(* IEC 61131-3 sources: volt/packages/volt-lsp-iec/test-corpus/bakon-nano/Device/Plc Logic/Application/Library Manager/AlarmManager (part 4) *)

(* ---- STANDARDALARMCONFIGURATION.pou ---- *)
FUNCTION_BLOCK STANDARDALARMCONFIGURATION
VAR
	M_PAITFALARMGROUPS : POINTER TO ARRAY [0..0] OF IAlarmGroup;
	M_ICOUNTALARMGROUPS : INT;
	M_PAITFALARMCLASSES : POINTER TO ARRAY [0..0] OF IAlarmClass;
	M_ICOUNTALARMCLASSES : INT;
	M_XVARIABLESREGISTERED : BOOL;
	M_XFIRST : BOOL;
	M_XPLACEHOLDANALYZED : BOOL;
	M_LTSTARTTIME : LTIME;
	M_DATABASESIZELIMIT : DatabaseSizeLimit;
	M_XDATABASESIZELIMITBLOCKED : BOOL;
	_XRAISEDMOREALARMSTHANSTORAGELIMITREPORTED : BOOL;
	_XCLEARHISTORY : BOOL;
	_XKEEPACTIVEALARMS : BOOL;
	M_DICTALARMTEMPLATEINSTANCES : AlarmInstanceDictionary;
	M_SZAPPNAME : STRING(CmpApp.GlobalConstants.MAX_LEN_APPLNAME);
	DATABASESIZELIMIT : IDatabaseSizeLimit;
	TOTALROWSTOINSERT : UDINT;
END_VAR
END_FUNCTION_BLOCK

METHOD FB_EXIT : BOOL
VAR_INPUT
	BINCOPYCODE : BOOL;
END_VAR
END_METHOD

METHOD FB_INIT : BOOL
VAR_INPUT
	BINITRETAINS : BOOL;
	BINCOPYCODE : BOOL;
END_VAR
END_METHOD

METHOD FINDALARMBYID : IAlarm
VAR_INPUT
	USIALARMGROUPID : ALARMGROUP_ID;
	UIALARMID : ALARM_ID;
END_VAR
END_METHOD

METHOD REGISTERVARIABLES
END_METHOD

METHOD ADDTOINSTANCEDICTIONARY : BOOL
VAR_INPUT
	PINSTANCE : POINTER TO BYTE;
	PSTALARMTEMPLATENAME : POINTER TO STRING;
	UDIALARMGROUPID : UDINT;
	UITEMPLATEALARMSOFFSET : UINT;
	UITEMPLATEALARMSLENGTH : UINT;
	UITEMPLATEEVENTSOFFSET : UINT;
	UITEMPLATEEVENTSLENGTH : UINT;
END_VAR
END_METHOD

METHOD CLEARINSTANCEDICTIONARY : BOOL
END_METHOD

METHOD GETALARMFROMDICTIONARY : IAlarm8
VAR_INPUT
	PINSTANCE : POINTER TO BYTE;
	UDIALARMID : REFERENCE TO ALARM_ID;
	STALARMTEMPLATENAME : REFERENCE TO STRING;
END_VAR
VAR_OUTPUT
	USIALARMGROUPID : ALARMGROUP_ID;
	UIALARMID : ALARM_ID;
END_VAR
END_METHOD

METHOD CREATEALARMSTORAGETASK
VAR_INPUT
	STSTORAGETASKGROUPNAME : REFERENCE TO STRING;
END_VAR
END_METHOD

METHOD INITSTORAGETASKINFO
VAR_INPUT
	ITASKPRIORITY : INT;
	DWINTERVAL : DWORD;
END_VAR
END_METHOD

METHOD ACKNOWLEDGEALL
END_METHOD

METHOD ACKNOWLEDGEALLOFGROUP
VAR_INPUT
	USIALARMGROUPID : ALARMGROUP_ID;
END_VAR
END_METHOD

METHOD ACKNOWLEDGEONEOFGROUP
VAR_INPUT
	USIALARMGROUPID : ALARMGROUP_ID;
	UIALARMID : ALARM_ID;
END_VAR
END_METHOD

METHOD CYCLICCALL
END_METHOD

METHOD FINDALARM : POINTER TO Alarm
VAR_INPUT
	SALARMGROUP : STRING;
	UIALARMID : ALARM_ID;
END_VAR
END_METHOD

METHOD FINDALARMCLASS : IAlarmClass
VAR_INPUT
	UDIID : UDINT;
END_VAR
END_METHOD

METHOD FINDALARMGROUP : IAlarmGroup
VAR_INPUT
	UDIID : UDINT;
END_VAR
END_METHOD

METHOD GETSTORAGE : IDatabaseFileAlarmStorage
END_METHOD

METHOD HASSTORAGE : BOOL
END_METHOD

METHOD RAISEEVENT : BOOL
VAR_INPUT
	EVENT : AlarmEvent;
END_VAR
END_METHOD

METHOD DETERMINERELEVANTALARMS : UDINT
VAR_INPUT
	ITFALARMFILTERCRITERIA : IAlarmFilterCriteria;
	PARRITFRELEVANTALARMS : POINTER TO ARRAY [0..0] OF IAlarm;
	IOFFSET : INT;
END_VAR
END_METHOD

METHOD FINDALARMGROUPBYNAME : IAlarmGroup
VAR_INPUT
	SALARMGROUP : STRING;
END_VAR
END_METHOD

METHOD FINDALARMCLASSBYNAME : IAlarmClass
VAR_INPUT
	SALARMCLASS : STRING;
END_VAR
END_METHOD

METHOD RAISEEVENT2 : BOOL
VAR_INPUT
	EVENT : AlarmEvent;
END_VAR
VAR_OUTPUT
	ITFALARM : IAlarm;
END_VAR
END_METHOD

METHOD GETALARMGROUPS : POINTER TO ARRAY [0..0] OF IAlarmGroup
VAR_OUTPUT
	IALARMGROUPCOUNT : INT;
END_VAR
END_METHOD

METHOD FINDALARMCLASSCOUNT : INT
END_METHOD

METHOD CLEARHISTORY : BOOL
VAR_INPUT
	XKEEPACTIVEALARMS : BOOL;
END_VAR
END_METHOD

METHOD ACKNOWLEDGEALLOFGROUPWITHCOMMENT
VAR_INPUT
	USIALARMGROUPID : ALARMGROUP_ID;
END_VAR
VAR_IN_OUT
	WSCOMMENT : WSTRING;
	WSUSERID : WSTRING;
END_VAR
END_METHOD

METHOD ACKNOWLEDGEALLWITHCOMMENT
VAR_IN_OUT
	WSCOMMENT : WSTRING;
	WSUSERID : WSTRING;
END_VAR
END_METHOD

METHOD ACKNOWLEDGEONEOFGROUPWITHCOMMENT
VAR_INPUT
	USIALARMGROUPID : ALARMGROUP_ID;
	UIALARMID : ALARM_ID;
END_VAR
VAR_IN_OUT
	WSCOMMENT : WSTRING;
	WSUSERID : WSTRING;
END_VAR
END_METHOD

METHOD SETCOMMENT : UDINT
VAR_INPUT
	USIALARMGROUPID : ALARMGROUP_ID;
	UIALARMID : ALARM_ID;
END_VAR
VAR_IN_OUT
	WSCOMMENT : WSTRING;
	WSUSERID : WSTRING;
END_VAR
END_METHOD

METHOD TRAVERSEALLALARMSOFALLALARMGROUPS
VAR_INPUT
	ITFALARMTRAVERSALCONSUMER : IAlarmTraversalConsumer;
END_VAR
END_METHOD

METHOD TRAVERSEALLCLASSES
VAR_INPUT
	ITFALARMTRAVERSALCONSUMER : IAlarmTraversalConsumer;
END_VAR
END_METHOD

METHOD NOTIFYREINITDONE
END_METHOD

METHOD CLEARALLALARMHISTORYENTRIESIFWISHED : BOOL
VAR_INPUT
	ITFDATABASEFILEALARMSTORAGE : IDatabaseFileAlarmStorage;
END_VAR
END_METHOD

METHOD CLEARONLYHISTORYOFINACTIVEALARMS : BOOL
END_METHOD

METHOD PRVACKNOWLEDGE
VAR_INPUT
	PAALARMS : POINTER TO ARRAY [0..0] OF Alarm;
	IALARMCOUNT : INT;
	UIALARMID : ALARM_ID;
	XACKALL : BOOL;
	PWSCOMMENT : POINTER TO WSTRING;
	PWSUSER : POINTER TO WSTRING;
END_VAR
END_METHOD

METHOD PRVCHECKSETACKNOWLEDGE
VAR_INPUT
	INDEX : INT;
	UIALARMID : ALARM_ID;
	XACKALL : BOOL;
	PWSCOMMENT : POINTER TO WSTRING;
	PWSUSER : POINTER TO WSTRING;
END_VAR
END_METHOD

METHOD PRVCREATEALARMSTORAGEMETADATAFILE
END_METHOD

METHOD PRVDETERMINERELEVANTALARMS : UDINT
VAR_INPUT
	PAALARMS : POINTER TO ARRAY [0..0] OF Alarm;
	IALARMCOUNT : INT;
	ITFALARMFILTERCRITERIA : IAlarmFilterCriteria;
	PARRITFRELEVANTALARMS : POINTER TO ARRAY [0..0] OF IAlarm;
	IOFFSET : INT;
END_VAR
END_METHOD

METHOD PRVINITIALIZEALARMCONFIGURATION
END_METHOD

METHOD PRVTRYGETCURRENTROW : BOOL
VAR_OUTPUT
	CURRENTROW : AlarmStorageRow;
END_VAR
END_METHOD

METHOD PRVTSTPLACEHOLDERS : BOOL
VAR_INPUT
	ALARM : REFERENCE TO Alarm;
END_VAR
END_METHOD

METHOD PRVWITHBRACKETS : STRING
VAR_INPUT
	SSTRING : STRING;
END_VAR
END_METHOD

METHOD PRVWITHOPENINGBRACKET : STRING
VAR_INPUT
	SSTRING : STRING;
END_VAR
END_METHOD

(* ---- STANDARDALARMCONFIGURATIONREMOTE.pou ---- *)
FUNCTION_BLOCK STANDARDALARMCONFIGURATIONREMOTE
VAR_INPUT
	M_PAITFPROXY : POINTER TO ARRAY [0..10] OF IProxy;
	M_IPROXYNUM : INT;
END_VAR
VAR
	M_SIALREADYSCAN : SINT := -1;
	PROXYNUM : INT;
END_VAR
END_FUNCTION_BLOCK

METHOD CYCLICCALL
END_METHOD

METHOD GETACTIVEALARMS
VAR_INPUT
	PASNAME : POINTER TO ARRAY [0..10] OF STRING;
	IGROUPCOUNT : INT;
	FILTERCRITERIA : REFERENCE TO VisuFbAlarmFilterCriteria;
	ITFALARMDATABLOCK : IAlarmDataBlockBaseDINT;
END_VAR
VAR_IN_OUT
	DISTUBPROG : DINT;
END_VAR
END_METHOD

METHOD GETALARMCLASSDESC : BOOL
VAR_INPUT
	SPROXYNAME : STRING;
	UDIID : UDINT;
END_VAR
VAR_OUTPUT
	SDESC : ProxyStructAlarmClassDesc;
END_VAR
END_METHOD

METHOD GETALARMCLASSDESCBYNAME : BOOL
VAR_INPUT
	SPROXYNAME : STRING;
	SCLASSNAME : STRING;
END_VAR
VAR_OUTPUT
	SDESC : ProxyStructAlarmClassDesc;
END_VAR
END_METHOD

METHOD GETALARMDESC : BOOL
VAR_INPUT
	SPROXYNAME : STRING;
	UDIALMID : UDINT;
	UDIGRPID : UDINT;
END_VAR
VAR_OUTPUT
	SDESC : ProxyStructAlarmDesc;
END_VAR
END_METHOD

METHOD GETALARMDISPLAYOPTIONS : BOOL
VAR_INPUT
	ITFALARMMETAOBJECTSTUB5 : IAlarmMetaObjectStub5;
	REFDISPLAYOPTIONS : REFERENCE TO DisplayOptions;
END_VAR
VAR_OUTPUT
	XVALID : BOOL;
	SCLASSREMAP : STRING;
END_VAR
END_METHOD

METHOD GETALARMGROUPDESC : BOOL
VAR_INPUT
	SPROXYNAME : STRING;
	UDIID : UDINT;
END_VAR
VAR_OUTPUT
	SDESC : ProxyStructAlarmGroupDesc;
END_VAR
END_METHOD

METHOD GETALARMGROUPDESCBYNAME : BOOL
VAR_INPUT
	SPROXYNAME : STRING;
	SGRPNAME : STRING;
END_VAR
VAR_OUTPUT
	SDESC : ProxyStructAlarmGroupDesc;
END_VAR
END_METHOD

METHOD GETALARMMESSAGE : BOOL
VAR_INPUT
	ITFALARMMETAOBJECTSTUB5 : IAlarmMetaObjectStub5;
	IWHICHMESSAGE : INT;
	REFCHARBUFFERSTRING : REFERENCE TO CharBufferString;
	STRINGTYPE : __SYSTEM.TYPE_CLASS;
END_VAR
END_METHOD

METHOD GETALARMMESSAGE2 : BOOL
VAR_INPUT
	SNAME : STRING;
	STEXTLISTNAME : STRING;
	STEXTLISTINDEX : STRING;
	IWHICHMESSAGE : INT;
	STRINGTYPE : __SYSTEM.TYPE_CLASS;
END_VAR
VAR_OUTPUT
	MESSAGE : CharBufferPtr;
END_VAR
END_METHOD

METHOD GETPROXY : IProxy
VAR_INPUT
	SNAME : STRING;
END_VAR
END_METHOD

METHOD GETSTORAGE : IDatabaseFileAlarmStorage
END_METHOD

METHOD HASSTORAGE : BOOL
END_METHOD

METHOD REGISTERUSERCLIENT : BOOL
VAR_INPUT
	IINDEX : INT;
END_VAR
VAR_OUTPUT
	ITFPROXY : IProxy;
END_VAR
END_METHOD

METHOD SETALARMSTOACK
VAR_INPUT
	ITFALARMDATABLOCK : IAlarmDataBlockBase2;
END_VAR
END_METHOD

METHOD REMOTEDEVICEREACHED
VAR_INPUT
	ROW : REFERENCE TO AlarmStorageRow;
	XFIRST : BOOL;
	IVERSION : INT;
END_VAR
END_METHOD

METHOD PRVGETPROXY : IProxy
VAR_INPUT
	SNAME : STRING;
END_VAR
END_METHOD

METHOD GETPROXYALARMCLASSESDESCRIPTION : BOOL
VAR_INPUT
	SNAME : STRING;
	PCLDESC : POINTER TO ARRAY [0..0] OF ProxyStructMonitorAlarmClassDesc;
	ISIZE : INT;
END_VAR
VAR_OUTPUT
	ICLCNT : INT;
END_VAR
END_METHOD

METHOD GETPROXYALARMGROUPSDESCRIPTION : BOOL
VAR_INPUT
	SNAME : STRING;
	PGRPDESC : POINTER TO ARRAY [0..0] OF ProxyStructMonitorAlarmGroupDesc;
	ISIZE : INT;
END_VAR
VAR_OUTPUT
	IGRPCNT : INT;
END_VAR
END_METHOD

METHOD GETPROXYALARMSDESCRIPTION : BOOL
VAR_INPUT
	SNAME : STRING;
	PALMDESC : POINTER TO ARRAY [0..0] OF ProxyStructMonitorAlarmDesc;
	DISIZE : DINT;
END_VAR
VAR_OUTPUT
	DIALMCNT : DINT;
END_VAR
END_METHOD

METHOD GETPROXYSTATISTICS : BOOL
VAR_INPUT
	SNAME : STRING;
END_VAR
VAR_OUTPUT
	STRUCTMONITOR : ProxyStructMonitor;
END_VAR
END_METHOD

METHOD GETPROXYSTATISTICSSINGLEACTIVITY : BOOL
VAR_INPUT
	SNAME : STRING;
	ITASKID : INT;
END_VAR
VAR_OUTPUT
	STRUCTMONITOR : ProxyStructMonitorRequest;
END_VAR
END_METHOD

(* ---- STANDARDALARMHANDLER.pou ---- *)
FUNCTION_BLOCK STANDARDALARMHANDLER
VAR
	M_AITFALARMCONFIGURATIONS : ARRAY [0..(MAX_COUNT_CONFIG - 1)] OF IAlarmConfiguration;
	M_ICOUNTCONFIGURATIONS : INT := 0;
	M_AITFALARMCONFIGURATIONSREM : ARRAY [0..(MAX_COUNT_CONFIG - 1)] OF IAlarmConfigurationRemote;
	M_ICOUNTCONFIGURATIONSREM : INT := 0;
	M_ALARMMANAGERCLIENTINFOSTRUCTVECTOR : AlarmManagerClientInfoStructVector;
	M_DIALARMSTATETRANSITIONCOUNTERPREVIOUSCALL : DINT;
	M_DIALARMSTORAGECOUNTERPREVIOUSCALL : DINT;
	M_ITFSTORAGETODELETE : IDatabaseFileAlarmStorage;
	M_XSTART : BOOL := TRUE;
	M_XFIRSTCYCLEAFTERDOWNLOAD : BOOL := TRUE;
	MAX_COUNT_CONFIG : BYTE := 2;
	ALARMCONFIGURATIONCOUNT : INT;
	ISREADY : BOOL;
END_VAR
END_FUNCTION_BLOCK

METHOD FB_EXIT : BOOL
VAR_INPUT
	BINCOPYCODE : BOOL;
END_VAR
END_METHOD

METHOD FB_INIT : BOOL
VAR_INPUT
	BINITRETAINS : BOOL;
	BINCOPYCODE : BOOL;
END_VAR
END_METHOD

METHOD FINDALARM : POINTER TO Alarm
VAR_INPUT
	SALARMGROUP : STRING;
	UIALARMID : ALARM_ID;
END_VAR
END_METHOD

METHOD FINDALARMCLASSBYNAME : IAlarmClass
VAR_INPUT
	SALARMCLASS : STRING;
END_VAR
END_METHOD

METHOD FINDALARMCLASSCOUNTALL : INT
END_METHOD

METHOD FINDALARMGROUPBYNAME : IAlarmGroup
VAR_INPUT
	SALARMGROUP : STRING;
END_VAR
END_METHOD

METHOD FINDALARMGROUPBYNAMEALL : IAlarmGroup
VAR_INPUT
	SALARMGROUP : STRING;
END_VAR
END_METHOD

METHOD REREGISTERCLIENTS
END_METHOD

METHOD TRAVERSEALLALARMSOFALLALARMCONFIGURATIONS
VAR_INPUT
	ITFALARMTRAVERSALCONSUMER : IAlarmTraversalConsumer;
END_VAR
END_METHOD

METHOD TRAVERSEALLCLASSESOFALLALARMCONFIGURATIONS
VAR_INPUT
	ITFALARMTRAVERSALCONSUMER : IAlarmTraversalConsumer;
END_VAR
END_METHOD

METHOD ALLOCBYTES : POINTER TO BYTE
VAR_INPUT
	UXISIZE : __UXINT;
END_VAR
END_METHOD

METHOD ALLOCFBALARMCLASSADAPTER : POINTER TO AlarmClassAdapter
END_METHOD

METHOD ALLOCFBALARMGROUPADAPTER : POINTER TO AlarmGroupAdapter
END_METHOD

METHOD ALLOCVALUETYPEBUNDLE : POINTER TO ValueTypeBundle
END_METHOD

METHOD ACKNOWLEDGEALL
END_METHOD

METHOD ACKNOWLEDGEALLOFGROUP
VAR_INPUT
	USIALARMGROUPID : ALARMGROUP_ID;
END_VAR
END_METHOD

METHOD ACKNOWLEDGEONEOFGROUP
VAR_INPUT
	USIALARMGROUPID : ALARMGROUP_ID;
	UIALARMID : ALARM_ID;
END_VAR
END_METHOD

METHOD CYCLICCALL
END_METHOD

METHOD FINDALARMCLASS : IAlarmClass
VAR_INPUT
	UDIID : UDINT;
END_VAR
END_METHOD

METHOD FINDALARMGROUP : IAlarmGroup
VAR_INPUT
	UDIID : UDINT;
END_VAR
END_METHOD

METHOD GETSTORAGE : IDatabaseFileAlarmStorage
END_METHOD

METHOD HASSTORAGE : BOOL
END_METHOD

METHOD RAISEEVENT : BOOL
VAR_INPUT
	USIALARMGROUPID : ALARMGROUP_ID;
	UIALARMID : ALARM_ID;
END_VAR
END_METHOD

METHOD REGISTERALARMCONFIGURATION
VAR_INPUT
	ITFALARMCONFIGURATION : IAlarmConfiguration;
END_VAR
END_METHOD

METHOD GETACTIVEALARMS : UDINT
VAR_INPUT
	ITFALARMMANAGERCLIENT : IAlarmManagerClient;
END_VAR
VAR_OUTPUT
	PARRITFACTIVEALARMS : POINTER TO ARRAY [0..0] OF IAlarm;
	ICOUNTACTIVEALARMS : INT;
END_VAR
END_METHOD

METHOD GETALARMSFROMSTORAGE : UDINT
VAR_INPUT
	ITFALARMMANAGERCLIENT : IAlarmManagerClient;
	ISKIPROWS : INT;
END_VAR
VAR_OUTPUT
	ICOUNTROWS : INT;
END_VAR
VAR_IN_OUT
	BROWIDVALID : BOOL;
	DIROWID : DINT;
END_VAR
END_METHOD

METHOD GETCOUNTALARMSFROMSTORAGE : DINT
VAR_INPUT
	ITFALARMMANAGERCLIENT : IAlarmManagerClient;
END_VAR
VAR_OUTPUT
	UDIRESULT : UDINT;
END_VAR
END_METHOD

METHOD REGISTERCLIENT : UDINT
VAR_INPUT
	ITFALARMMANAGERCLIENT : IAlarmManagerClient;
	PARRITFALARMSFROMHISTORY : POINTER TO ARRAY [0..0] OF IAlarm2;
	ICOUNTALARMSFROMHISTORY : INT;
END_VAR
END_METHOD

METHOD UNREGISTERCLIENT : UDINT
VAR_INPUT
	ITFALARMMANAGERCLIENT : IAlarmManagerClient;
END_VAR
END_METHOD

METHOD UNREGISTERALARMCONFIGURATION
VAR_INPUT
	ITFALARMCONFIGURATION : IAlarmConfiguration;
END_VAR
END_METHOD

METHOD REGISTERALARMSTATECHANGEDLISTENER : BOOL
VAR_INPUT
	ITFALARMSTATECHANGEDLISTENER : IAlarmStateChangedListener;
END_VAR
END_METHOD

METHOD GETALARMCONFIGURATION : IAlarmConfiguration
VAR_INPUT
	IPOS : INT;
END_VAR
END_METHOD

METHOD ACKNOWLEDGEALLOFGROUPWITHCOMMENT
VAR_INPUT
	USIALARMGROUPID : ALARMGROUP_ID;
END_VAR
VAR_IN_OUT
	WSCOMMENT : WSTRING;
	WSUSERID : WSTRING;
END_VAR
END_METHOD

METHOD ACKNOWLEDGEALLWITHCOMMENT
VAR_IN_OUT
	WSCOMMENT : WSTRING;
	WSUSERID : WSTRING;
END_VAR
END_METHOD

METHOD ACKNOWLEDGEONEOFGROUPWITHCOMMENT
VAR_INPUT
	USIALARMGROUPID : ALARMGROUP_ID;
	UIALARMID : ALARM_ID;
END_VAR
VAR_IN_OUT
	WSCOMMENT : WSTRING;
	WSUSERID : WSTRING;
END_VAR
END_METHOD

METHOD SETCOMMENT : UDINT
VAR_INPUT
	USIALARMGROUPID : ALARMGROUP_ID;
	UIALARMID : ALARM_ID;
END_VAR
VAR_IN_OUT
	WSCOMMENT : WSTRING;
	WSUSERID : WSTRING;
END_VAR
END_METHOD

METHOD GETINSTANCEALARM : IAlarm8
VAR_INPUT
	PFBINSTANCE : POINTER TO BYTE;
	UITEMPLATEALARMID : ALARM_ID;
END_VAR
VAR_OUTPUT
	USIALARMGROUPID : ALARMGROUP_ID;
	UIALARMID : ALARM_ID;
END_VAR
END_METHOD

METHOD GETINSTANCEALARMBYNAME : IAlarm8
VAR_INPUT
	PFBINSTANCE : POINTER TO BYTE;
	UITEMPLATEALARMID : ALARM_ID;
	STALARMTEMPLATENAME : STRING(255);
END_VAR
VAR_OUTPUT
	USIALARMGROUPID : ALARMGROUP_ID;
	UIALARMID : ALARM_ID;
END_VAR
END_METHOD

METHOD RAISEEVENTALARMINSTANCE : BOOL
VAR_INPUT
	PFBINSTANCE : POINTER TO BYTE;
	UITEMPLATEALARMID : ALARM_ID;
END_VAR
END_METHOD

METHOD RAISEEVENTALARMINSTANCEBYNAME : BOOL
VAR_INPUT
	PFBINSTANCE : POINTER TO BYTE;
	UITEMPLATEALARMID : ALARM_ID;
	STALARMTEMPLATENAME : STRING(255);
END_VAR
END_METHOD

METHOD ACTIVATEALARM : BOOL
VAR_INPUT
	USIALARMGROUPID : ALARMGROUP_ID;
	UIALARMID : ALARM_ID;
END_VAR
END_METHOD

METHOD ACTIVATEALARMINSTANCE : BOOL
VAR_INPUT
	PFBINSTANCE : POINTER TO BYTE;
	UITEMPLATEALARMID : ALARM_ID;
END_VAR
END_METHOD

METHOD DEACTIVATEALARM : BOOL
VAR_INPUT
	USIALARMGROUPID : ALARMGROUP_ID;
	UIALARMID : ALARM_ID;
END_VAR
END_METHOD

METHOD DEACTIVATEALARMINSTANCE : BOOL
VAR_INPUT
	PFBINSTANCE : POINTER TO BYTE;
	UITEMPLATEALARMID : ALARM_ID;
END_VAR
END_METHOD

METHOD GETALARMIDANDALARMGROUPNAME : BOOL
VAR_INPUT
	UDIALARMGROUPID : UDINT;
	UDIALARMID : UDINT;
END_VAR
VAR_OUTPUT
	SALARMGROUPNAME : STRING;
	UIALARMID : ALARM_ID;
END_VAR
END_METHOD

METHOD GETACTIVEALARMSFROMPROXY
VAR_INPUT
	PASNAME : POINTER TO ARRAY [0..10] OF STRING;
	IGROUPCOUNT : INT;
	FILTERCRITERIA : REFERENCE TO VisuFbAlarmFilterCriteria;
	ITFALARMDATABLOCK : IAlarmDataBlockBaseDINT;
END_VAR
VAR_IN_OUT
	DISTUBPROG : DINT;
END_VAR
END_METHOD

METHOD GETALARMCLASSDESCBYNAMEFROMPROXY
VAR_INPUT
	SPROXYNAME : STRING;
	SCLASSNAME : STRING;
END_VAR
VAR_OUTPUT
	SDESC : ProxyStructAlarmClassDesc;
END_VAR
END_METHOD

METHOD GETALARMCLASSDESCFROMPROXY
VAR_INPUT
	SNAME : STRING;
	UDIID : UDINT;
END_VAR
VAR_OUTPUT
	SDESC : ProxyStructAlarmClassDesc;
END_VAR
END_METHOD

METHOD GETALARMDESCFROMPROXY
VAR_INPUT
	SNAME : STRING;
	UDIALMID : UDINT;
	UDIGRPID : UDINT;
END_VAR
VAR_OUTPUT
	SDESC : ProxyStructAlarmDesc;
END_VAR
END_METHOD

METHOD GETALARMDISPLAYOPTIONSFROMPROXY
VAR_INPUT
	ITFALARMMETAOBJECTSTUB5 : IAlarmMetaObjectStub5;
	REFDISPLAYOPTIONS : REFERENCE TO DisplayOptions;
END_VAR
VAR_OUTPUT
	XVALID : BOOL;
	SCLASSREMAP : STRING;
END_VAR
END_METHOD

METHOD GETALARMGROUPDESCBYNAMEFROMPROXY
VAR_INPUT
	SPROXYNAME : STRING;
	SGRPNAME : STRING;
END_VAR
VAR_OUTPUT
	SDESC : ProxyStructAlarmGroupDesc;
END_VAR
END_METHOD

METHOD GETALARMGROUPDESCFROMPROXY
VAR_INPUT
	SNAME : STRING;
	UDIID : UDINT;
END_VAR
VAR_OUTPUT
	SDESC : ProxyStructAlarmGroupDesc;
END_VAR
END_METHOD

METHOD GETALARMMESSAGEFROMPROXY
VAR_INPUT
	ITFALARMMETAOBJECTSTUB5 : IAlarmMetaObjectStub5;
	IWHICHMESSAGE : INT;
	REFCHARBUFFERSTRING : REFERENCE TO CharBufferString;
	STRINGTYPE : __SYSTEM.TYPE_CLASS;
END_VAR
END_METHOD

METHOD GETALARMMESSAGEFROMPROXY2
VAR_INPUT
	SNAME : STRING;
	STEXTLISTNAME : STRING;
	STEXTLISTINDEX : STRING;
	IWHICHMESSAGE : INT;
	STRINGTYPE : __SYSTEM.TYPE_CLASS;
END_VAR
VAR_OUTPUT
	MESSAGE : CharBufferPtr;
END_VAR
END_METHOD

METHOD GETPROXY : IProxy
VAR_INPUT
	SNAME : STRING;
END_VAR
END_METHOD

METHOD REGISTERALARMCONFIGURATIONREMOTE
VAR_INPUT
	ITFALARMCONFIGURATION : IAlarmConfigurationRemote;
END_VAR
END_METHOD

METHOD SETALARMSTOACKPROXY
VAR_INPUT
	ITFALARMDATABLOCK : IAlarmDataBlockBase2;
END_VAR
END_METHOD

METHOD GETPROXYALARMCLASSESDESCRIPTION : BOOL
VAR_INPUT
	SNAME : STRING;
	PCLDESC : POINTER TO ARRAY [0..0] OF ProxyStructMonitorAlarmClassDesc;
	ISIZE : INT;
END_VAR
VAR_OUTPUT
	ICLCNT : INT;
END_VAR
END_METHOD

METHOD GETPROXYALARMGROUPSDESCRIPTION : BOOL
VAR_INPUT
	SNAME : STRING;
	PGRPDESC : POINTER TO ARRAY [0..0] OF ProxyStructMonitorAlarmGroupDesc;
	ISIZE : INT;
END_VAR
VAR_OUTPUT
	IGRPCNT : INT;
END_VAR
END_METHOD

METHOD GETPROXYALARMSDESCRIPTION : BOOL
VAR_INPUT
	SNAME : STRING;
	PALMDESC : POINTER TO ARRAY [0..0] OF ProxyStructMonitorAlarmDesc;
	DISIZE : DINT;
END_VAR
VAR_OUTPUT
	DIALMCNT : DINT;
END_VAR
END_METHOD

METHOD GETPROXYSTATISTICS : BOOL
VAR_INPUT
	SNAME : STRING;
END_VAR
VAR_OUTPUT
	STRUCTMONITOR : ProxyStructMonitor;
END_VAR
END_METHOD

METHOD GETPROXYSTATISTICSSINGLEACTIVITY : BOOL
VAR_INPUT
	SNAME : STRING;
	ITASKID : INT;
END_VAR
VAR_OUTPUT
	STRUCTMONITOR : ProxyStructMonitorRequest;
END_VAR
END_METHOD

METHOD CLEARTEMPLATEDICTIONARY : BOOL
END_METHOD

METHOD REGISTERTEMPLATEINSTANCE : BOOL
VAR_INPUT
	PINSTANCE : POINTER TO BYTE;
	UDIALARMGROUPID : UDINT;
	UITEMPLATEALARMSOFFSET : UINT;
	UITEMPLATEALARMSLENGTH : UINT;
	PSTALARMTEMPLATENAME : POINTER TO STRING;
	UITEMPLATEEVENTSOFFSET : UINT;
	UITEMPLATEEVENTSLENGTH : UINT;
END_VAR
END_METHOD

METHOD INITAFTERDOWNLOAD : BOOL
END_METHOD

METHOD PRVCHECKALARMMANAGERCLIENT : UDINT
VAR_INPUT
	ITFALARMMANAGERCLIENT : IAlarmManagerClient;
END_VAR
END_METHOD

METHOD PRVCHECKVALIDEVENT : BOOL
VAR_IN_OUT
	UIALARMID : ALARM_ID;
	PALARM8 : IAlarm8;
END_VAR
END_METHOD

METHOD PRVFREECLIENT : UDINT
VAR_INPUT
	PALARMMANAGERCLIENTINFOSTRUCT : POINTER TO AlarmManagerClientInfoStruct;
END_VAR
END_METHOD

METHOD PRVNOTIFYALARMMANAGERCLIENT
VAR_INPUT
	ITFALARMMANAGERCLIENT : IAlarmManagerClient;
	ITFALARM4 : IAlarm4;
END_VAR
END_METHOD

(* ---- STATECOMPARER.pou ---- *)
FUNCTION_BLOCK STATECOMPARER EXTENDS TSLastComparer
END_FUNCTION_BLOCK

METHOD COMPARE : INT
VAR_INPUT
	DIINDEXALARM1 : DINT;
	DIINDEXALARM2 : DINT;
END_VAR
END_METHOD

(* ---- STATISTICS_LTIME.pou ---- *)
FUNCTION_BLOCK STATISTICS_LTIME
VAR_INPUT
	XENABLE : BOOL;
	LTINPUT : LTIME;
END_VAR
VAR
	LTMIN : LTIME;
	LTMAX : LTIME;
	LTAVERAGE : LTIME;
	LICOUNTER : LINT;
	LISUM : LINT;
	XOLDENABLE : BOOL;
	LIAVERAGE : LINT;
	AVERAGE : LTIME;
	COUNT : LINT;
	MAXIMUM : LTIME;
	MINIMUM : LTIME;
END_VAR
END_FUNCTION_BLOCK

(* ---- STRINGCONTAINER.pou ---- *)
FUNCTION_BLOCK STRINGCONTAINER
VAR
	M_BUFFERVECTOR : StringContainerBufferVector;
	M_UDINEXTALLOCATIONSIZE : UDINT := INITIAL_BUFFER_SIZE;
	COMPONENT : STRING := 'StringContainer';
	STRINGTYPE_STRING : UINT := 16;
	STRINGTYPE_WSTRING : UINT := 17;
	INITIAL_BUFFER_SIZE : UDINT := 512;
END_VAR
END_FUNCTION_BLOCK

METHOD ADDSTRING : CharBufferPtr
VAR_INPUT
	CBPMESSAGE : CharBufferPtr;
	TYPECLASS : __SYSTEM.TYPE_CLASS;
END_VAR
VAR_OUTPUT
	UDIERROR : UDINT;
	DISTRINGLENGTH : DINT;
END_VAR
END_METHOD

METHOD FB_EXIT : BOOL
VAR_INPUT
	BINCOPYCODE : BOOL;
END_VAR
END_METHOD

METHOD PRVALLOCATEBUFFER : UDINT
END_METHOD

METHOD PRVALLOCATEBUFFERIFNEEDED : UDINT
END_METHOD

METHOD PRVFINDSTRINGINBUFFER : POINTER TO BYTE
VAR_INPUT
	CBPMESSAGE : CharBufferPtr;
	TYPECLASS : __SYSTEM.TYPE_CLASS;
	UDIWHICHBUFFER : UDINT;
END_VAR
VAR_OUTPUT
	XFOUND : BOOL;
END_VAR
END_METHOD

METHOD PRVHASFREECAPACITY : BOOL
VAR_INPUT
	DICOUNTBYTESREQUIRED : DINT;
	UDIWHICHBUFFER : UDINT;
END_VAR
END_METHOD

METHOD PRVOPENBUFFER : StringContainerBufferInfo
VAR_INPUT
	UDIWHICHBUFFER : UDINT;
END_VAR
END_METHOD

METHOD PRVSTORESTRINGINBUFFER : POINTER TO BYTE
VAR_INPUT
	CBPMESSAGE : CharBufferPtr;
	UISTRINGTYPE : UINT;
	DICOUNTBYTESTOCOPY : DINT;
	DICOUNTBYTESFORSTRING : DINT;
	UDIWHICHBUFFER : UDINT;
END_VAR
END_METHOD

(* ---- STRINGCONTAINERBUFFERVECTOR.pou ---- *)
FUNCTION_BLOCK STRINGCONTAINERBUFFERVECTOR EXTENDS BaseVector
VAR
	_PAPBYSTRINGCONTAINERBUFFERS : POINTER TO ARRAY [0..MAX_NUM_ENTRIES] OF POINTER TO BYTE;
	MAX_NUM_ENTRIES : INT := 10;
END_VAR
END_FUNCTION_BLOCK

METHOD ADDSTRINGCONTAINERBUFFER : UDINT
VAR_INPUT
	PBYBUFFER : POINTER TO BYTE;
END_VAR
END_METHOD

METHOD GETSTRINGCONTAINERBUFFERAT : POINTER TO BYTE
VAR_INPUT
	UDIINDEX : UDINT;
END_VAR
VAR_OUTPUT
	UDIRESULT : UDINT;
END_VAR
END_METHOD

METHOD ABSTRASSIGN : UDINT
VAR_INPUT
	PBT : POINTER TO BYTE;
	UDIINDEX : UDINT;
END_VAR
END_METHOD

METHOD ABSTRDATAPTRCHANGED : UDINT
END_METHOD

METHOD ABSTRSIZEOFELEMENT : UDINT
END_METHOD

(* ---- TEXTHELPER.pou ---- *)
FUNCTION_BLOCK TEXTHELPER
VAR_OUTPUT
	TEXT : STO.TEXT;
END_VAR
END_FUNCTION_BLOCK

METHOD FB_EXIT : BOOL
VAR_INPUT
	BINCOPYCODE : BOOL;
END_VAR
END_METHOD

METHOD FROMSTRING : STO.ERROR
VAR_INPUT
	PS : POINTER TO STRING;
	FUNCTIONCALLER : INT;
END_VAR
END_METHOD

METHOD FROMWSTRING : STO.ERROR
VAR_INPUT
	PWS : POINTER TO WSTRING;
	FUNCTIONCALLER : INT;
END_VAR
END_METHOD

METHOD RELEASE
END_METHOD

(* ---- TIMESTAMPANDVALUESCONTAINER.pou ---- *)
FUNCTION_BLOCK TIMESTAMPANDVALUESCONTAINER
VAR
	M_LITIMESTAMPLAST : AlarmManager_Interfaces.Timestamp;
	M_LITIMESTAMPACTIVE : AlarmManager_Interfaces.Timestamp;
	M_LITIMESTAMPINACTIVE : AlarmManager_Interfaces.Timestamp;
	M_LITIMESTAMPACKNOWLEDGE : AlarmManager_Interfaces.Timestamp;
	M_TRIGGERVALUE : ValueTypeBundle;
	M_ALATCHVARIABLES : ARRAY [1..COUNT_LATCH_VARIABLES] OF ValueTypeBundle;
	COUNT_LATCH_VARIABLES : INT := 10;
END_VAR
END_FUNCTION_BLOCK

METHOD FILL : BOOL
VAR_INPUT
	ITFRANDOMALARMREADACCESS : IRandomAlarmReadAccess;
	DIINDEXALARM : DINT;
	ICOUNTLATCHVARIABLES : INT;
END_VAR
END_METHOD

METHOD GETCOUNTLATCHVARIABLES : USINT
END_METHOD

METHOD GETLATCHVARVALUE : AlarmManagerInternal_Interfaces.ITypedValue2
VAR_INPUT
	IWHICHLATCHVAR : INT;
END_VAR
END_METHOD

METHOD GETCURRENTVALUE : AlarmManagerInternal_Interfaces.ITypedValue
END_METHOD

METHOD GETLATCHVAR1VALUE : AlarmManager_Interfaces.ITypedValue
END_METHOD

METHOD GETLATCHVAR2VALUE : AlarmManager_Interfaces.ITypedValue
END_METHOD

METHOD GETTIMESTAMPACKNOWLEDGE : AlarmManager_Interfaces.Timestamp
END_METHOD

METHOD GETTIMESTAMPACTIVE : AlarmManager_Interfaces.Timestamp
END_METHOD

METHOD GETTIMESTAMPINACTIVE : AlarmManager_Interfaces.Timestamp
END_METHOD

METHOD GETTIMESTAMPLAST : AlarmManager_Interfaces.Timestamp
END_METHOD

METHOD GETTRIGGERVALUE : AlarmManager_Interfaces.ITypedValue
END_METHOD

METHOD GETALARMGROUP : STRING
END_METHOD

METHOD GETCHECKSUM : UDINT
END_METHOD

METHOD GETID : AlarmManager_Interfaces.ALARM_ID
END_METHOD

METHOD GETSTATE : INT
END_METHOD

METHOD SETACKNOWLEDGE
VAR_INPUT
	BACKNOWLEDGEMULTIPLE : BOOL;
END_VAR
END_METHOD

METHOD SETALARMGROUP
VAR_INPUT
	SALARMGROUP : STRING;
END_VAR
END_METHOD

METHOD SETID
VAR_INPUT
	UIID : AlarmManager_Interfaces.ALARM_ID;
END_VAR
END_METHOD

METHOD SETLATCHVAR1VALUE
VAR_INPUT
	ITFTYPEDVALUELATCHVAR1 : AlarmManager_Interfaces.ITypedValue;
END_VAR
END_METHOD

METHOD SETLATCHVAR2VALUE
VAR_INPUT
	ITFTYPEDVALUELATCHVAR2 : AlarmManager_Interfaces.ITypedValue;
END_VAR
END_METHOD

METHOD SETLATCHVARVALUE
VAR_INPUT
	IWHICHLATCHVAR : INT;
	ITFTYPEDVALUELATCHVAR : AlarmManagerInternal_Interfaces.ITypedValue;
END_VAR
END_METHOD

METHOD SETSTATE
VAR_INPUT
	ISTATE : INT;
END_VAR
END_METHOD

METHOD SETTIMESTAMPACKNOWLEDGE
VAR_INPUT
	LITIMESTAMPACKNOWLEDGE : AlarmManager_Interfaces.Timestamp;
END_VAR
END_METHOD

METHOD SETTIMESTAMPACTIVE
VAR_INPUT
	LITIMESTAMPACTIVE : AlarmManager_Interfaces.Timestamp;
END_VAR
END_METHOD

METHOD SETTIMESTAMPINACTIVE
VAR_INPUT
	LITIMESTAMPINACTIVE : AlarmManager_Interfaces.Timestamp;
END_VAR
END_METHOD

METHOD SETTIMESTAMPLAST
VAR_INPUT
	LITIMESTAMPLAST : AlarmManager_Interfaces.Timestamp;
END_VAR
END_METHOD

METHOD SETTRIGGERVALUE
VAR_INPUT
	ITFTYPEDVALUETRIGGER : AlarmManager_Interfaces.ITypedValue;
END_VAR
END_METHOD

(* ---- TL_ALARMSTATUS.pou ---- *)
FUNCTION_BLOCK TL_ALARMSTATUS
VAR
	M_TEXTLISTFILE : STRING(255);
	_STNAMESPACE : STRING;
END_VAR
END_FUNCTION_BLOCK

(* ---- TSACKCOMPARER.pou ---- *)
FUNCTION_BLOCK TSACKCOMPARER EXTENDS AbstractTimestampComparer
END_FUNCTION_BLOCK

METHOD PROTGETTIMESTAMP : BOOL
VAR_INPUT
	DIINDEXALARM : DINT;
END_VAR
VAR_OUTPUT
	LITIMESTAMP : TIMESTAMP;
END_VAR
END_METHOD

(* ---- TSACTIVECOMPARER.pou ---- *)
FUNCTION_BLOCK TSACTIVECOMPARER EXTENDS AbstractTimestampComparer
END_FUNCTION_BLOCK

METHOD PROTGETTIMESTAMP : BOOL
VAR_INPUT
	DIINDEXALARM : DINT;
END_VAR
VAR_OUTPUT
	LITIMESTAMP : TIMESTAMP;
END_VAR
END_METHOD

(* ---- TSINACTIVECOMPARER.pou ---- *)
FUNCTION_BLOCK TSINACTIVECOMPARER EXTENDS AbstractTimestampComparer
END_FUNCTION_BLOCK

METHOD PROTGETTIMESTAMP : BOOL
VAR_INPUT
	DIINDEXALARM : DINT;
END_VAR
VAR_OUTPUT
	LITIMESTAMP : TIMESTAMP;
END_VAR
END_METHOD

(* ---- TSLASTCOMPARER.pou ---- *)
FUNCTION_BLOCK TSLASTCOMPARER EXTENDS AbstractTimestampComparer
END_FUNCTION_BLOCK

METHOD PROTGETTIMESTAMP : BOOL
VAR_INPUT
	DIINDEXALARM : DINT;
END_VAR
VAR_OUTPUT
	LITIMESTAMP : TIMESTAMP;
END_VAR
END_METHOD

(* ---- TYPEDVALUEFORMATTER.pou ---- *)
FUNCTION_BLOCK TYPEDVALUEFORMATTER
VAR
	M_CBSSTRINGFORMATSTRINGINT : CharBufferString;
	M_CBSSTRINGFORMATSTRINGLONG : CharBufferString;
	M_CBSSTRINGFORMATSTRINGFLOAT : CharBufferString;
	M_CBSSTRINGFORMATSTRINGSTRING : CharBufferString;
	M_CBSSTRINGFORMATSTRINGWSTRING : CharBufferString;
	M_CBSWSTRINGFORMATSTRINGINT : CharBufferString;
	M_CBSWSTRINGFORMATSTRINGLONG : CharBufferString;
	M_CBSWSTRINGFORMATSTRINGFLOAT : CharBufferString;
	M_CBSWSTRINGFORMATSTRINGSTRING : CharBufferString;
	M_CBSWSTRINGFORMATSTRINGWSTRING : CharBufferString;
	M_APSTRINGFORMATSTRINGS : ARRAY [AlarmConstants.FMT_FIRST_FORMAT_STRING..AlarmConstants.FMT_LAST_FORMAT_STRING] OF POINTER TO CharBufferString;
	M_APWSTRINGFORMATSTRINGS : ARRAY [AlarmConstants.FMT_FIRST_FORMAT_STRING..AlarmConstants.FMT_LAST_FORMAT_STRING] OF POINTER TO CharBufferString;
END_VAR
END_FUNCTION_BLOCK

METHOD FB_EXIT : BOOL
VAR_INPUT
	BINCOPYCODE : BOOL;
END_VAR
END_METHOD

METHOD FB_INIT : BOOL
VAR_INPUT
	BINITRETAINS : BOOL;
	BINCOPYCODE : BOOL;
END_VAR
END_METHOD

METHOD FORMATTYPEDVALUE2 : CharBufferPtr
VAR_INPUT
	ITFTYPEDVALUE : ITypedValue;
	CBSRESULT : REFERENCE TO CharBufferString;
END_VAR
END_METHOD

(* ---- USERIDCOMPARER.pou ---- *)
FUNCTION_BLOCK USERIDCOMPARER EXTENDS TSLastComparer
END_FUNCTION_BLOCK

METHOD COMPARE : INT
VAR_INPUT
	DIINDEXALARM1 : DINT;
	DIINDEXALARM2 : DINT;
END_VAR
END_METHOD

(* ---- VALUECOMPARER.pou ---- *)
FUNCTION_BLOCK VALUECOMPARER EXTENDS TSLastComparer
VAR
	M_IWHICHVALUE : INT;
END_VAR
END_FUNCTION_BLOCK

METHOD BEFORECOMPARE
VAR_INPUT
	IWHICHVALUE : INT;
END_VAR
END_METHOD

METHOD COMPARE : INT
VAR_INPUT
	DIINDEXALARM1 : DINT;
	DIINDEXALARM2 : DINT;
END_VAR
END_METHOD

METHOD PRVCOMPARETYPE : INT
VAR_INPUT
	BYTYPE1 : BYTE;
	BYTYPE2 : BYTE;
END_VAR
VAR_OUTPUT
	ECOMPARABLETYPEBOTH : EComparableType;
	ENUMERIKCOMPARISON : ENumericComparison;
END_VAR
END_METHOD

METHOD PRVCOMPAREVALUE : INT
VAR_INPUT
	LIVALUE1 : LINT;
	BYTYPE1 : BYTE;
	LIVALUE2 : LINT;
	BYTYPE2 : BYTE;
	ECOMPARABLETYPEBOTH : EComparableType;
	ENUMERIKCOMPARISON : ENumericComparison;
END_VAR
END_METHOD

METHOD PRVCONVERTVALUETOLINT : LINT
VAR_INPUT
	LIVALUE : LINT;
	ITYPE : TypeClass;
END_VAR
END_METHOD

METHOD PRVGETCOMPARABLETYPE : EComparableType
VAR_INPUT
	BYTYPE : BYTE;
END_VAR
VAR_OUTPUT
	XISINT : BOOL;
	XISREAL : BOOL;
	XISLREAL : BOOL;
END_VAR
END_METHOD

METHOD PRVGETTYPE : BOOL
VAR_INPUT
	DIINDEXALARM : DINT;
END_VAR
VAR_OUTPUT
	BYTYPE : BYTE;
END_VAR
END_METHOD

METHOD PRVGETVALUE : BOOL
VAR_INPUT
	DIINDEXALARM : DINT;
END_VAR
VAR_OUTPUT
	LIVALUE : LINT;
END_VAR
END_METHOD

(* ---- VALUETYPEBUNDLE.pou ---- *)
FUNCTION_BLOCK VALUETYPEBUNDLE
VAR
	M_VALUE : ScalarType;
	M_TYPE : __SYSTEM.TYPE_CLASS := __SYSTEM.TYPE_CLASS.TYPE_NONE;
	M_ISTRINGSIZE : INT;
	M_PSSTRING : POINTER TO STRING(255);
	M_PWSSTRING : POINTER TO WSTRING(255);
END_VAR
END_FUNCTION_BLOCK

METHOD GETSIZE : INT
END_METHOD

METHOD GETTYPE : __SYSTEM.TYPE_CLASS
END_METHOD

METHOD GETVALUE : POINTER TO BYTE
END_METHOD

METHOD SETRAWVALUE
VAR_INPUT
	PABYVALUE : POINTER TO ARRAY [0..7] OF BYTE;
	ETYPETOSET : __SYSTEM.TYPE_CLASS;
END_VAR
END_METHOD

METHOD SETSTRINGSIZE
VAR_INPUT
	ISTRINGSIZE : INT;
END_VAR
END_METHOD

METHOD SETTYPE
VAR_INPUT
	TYPETOSET : __SYSTEM.TYPE_CLASS;
END_VAR
END_METHOD

METHOD SETVALUE
VAR_INPUT
	LIVALUE : LINT;
END_VAR
END_METHOD

(* ---- VISUFBALARMFILTERCRITERIA.pou ---- *)
FUNCTION_BLOCK VISUFBALARMFILTERCRITERIA
VAR_INPUT
	M_PSTARRALARMGROUPS : POINTER TO ARRAY [0..0] OF UDINT;
	M_ICOUNTALARMGROUPS : INT;
	M_BALLALARMGROUPS : BOOL;
	M_PSTARRALARMCLASSES : POINTER TO ARRAY [0..0] OF UDINT;
	M_ICOUNTALARMCLASSES : INT;
	M_BALLALARMCLASSES : BOOL;
	M_USIPRIORITYFROM : USINT;
	M_USIPRIORITYTO : USINT;
	M_PLATCH1VARIABLE : POINTER TO BYTE;
	M_ELATCH1VARTYPE : Visu_Types;
	M_PFILTTYPEVARIABLE : POINTER TO DWORD;
	M_DWFILTTYPEVARTYPE : DWORD;
	M_PDTFILTFROMVAR : POINTER TO DATE_AND_TIME;
	M_PDTFILTTOVAR : POINTER TO DATE_AND_TIME;
	M_PFILTTRTYPE : POINTER TO DWORD;
	M_DWFILTTRTYPE : DWORD;
	M_PARRALARMGROUPSREM : POINTER TO ARRAY [0..10] OF StruFilterRemoteAlm;
	M_ICOUNTALARMGROUPSREM : INT;
	M_BALLALARMGROUPSREM : BOOL;
	M_PARRALARMCLASSESREM : POINTER TO ARRAY [0..10] OF StruFilterRemoteAlm;
	M_ICOUNTALARMCLASSESREM : INT;
	M_BALLALARMCLASSESREM : BOOL;
	M_XFILTERLATCHAVAILABLE : BOOL;
	M_XFILTERTIMERANGEAVAILABLE : BOOL;
	M_EFILTERLATCHCONTENT : EFilterLatchContent;
	M_CRITERIA_LIFILTERCRITERIONTOSEARCH : LINT;
	M_CRITERIA_WVARIABLETYPETOSEARCH : WORD;
	M_CRITERIA_XVALIDSEARCH : BOOL;
	M_CRITERIA_XINDEX : BOOL;
END_VAR
VAR
	_FILTERLATCHCONTENT : EFilterLatchContent := EFilterLatchContent.NOT_SET;
	_VTYPE : Visu_Types;
	_LIVALUE : LINT;
	_RVALUE : REAL;
	_LRVALUE : LREAL;
	_PWSVALUE : POINTER TO WSTRING;
	_WSSTRVALUE : WSTRING(255);
	OLDIECSTRING : STRING(255);
	_FILTERTRTYPE : EFilterTimeRangeType := EFilterTimeRangeType.NOT_SET;
	_TSFROMVALUE : Timestamp;
	_TSTOVALUE : Timestamp;
	CNVIECTYPEDLITERAL : ConvertIecTypedLiteral;
	DWREASONNOTINDEX : DWORD;
	DWREASONNOTINDEXDISPLAYED : DWORD;
	XDISPTYPNOTCORRECT : BOOL;
	WOLDCHECKSUM : WORD;
	XDISPTSNOTCORRECT : BOOL;
	ERROR_FILTER_MASK_COMPILE : DWORD := 16#1;
	ERROR_FILTER_MASK_DISABLE : DWORD := 16#2;
	ERROR_FILTER_MASK_DB_OLD : DWORD := 16#4;
	ERROR_FILTER_MASK_SORT : DWORD := 16#8;
	ERROR_FILTER_MASK_DB_NOT_INDEXABLE : DWORD := 16#10;
	FILTERLATCHCONTENT : EFilterLatchContent;
	FILTERLATCHCONTENTASINT : INT;
	FILTERTIMERANGETYPE : EFilterTimeRangeType;
	FROMVALUELI : LINT;
	TOVALUELI : LINT;
	TYPEDLITERALTYPE : Visu_Types;
	VALUELI : LINT;
	VALUELREAL : LREAL;
	VALUEREAL : REAL;
	VALUEWSTRING : WSTRING;
	VALUEWSTRINGPOINTER : POINTER TO WSTRING;
END_VAR
END_FUNCTION_BLOCK

METHOD INITIALIZE
VAR_INPUT
	ITFALARMFILTERCRITERIA : IAlarmFilterCriteria;
END_VAR
END_METHOD

METHOD INITIALIZETODEFAULT
END_METHOD

METHOD ISFILTERCRITERIACHANGED : BOOL
END_METHOD

METHOD ISRELEVANTALARM : BOOL
VAR_INPUT
	ITFDATABASEACCESS : IDatabaseAccess;
	XREMOTEALM : BOOL;
	SPROXYNAME : STRING;
END_VAR
VAR_OUTPUT
	UDIGROUP : UDINT;
	BENDOFSEARCH : BOOL;
END_VAR
END_METHOD

METHOD MATCHESFILTERCRITERIA : BOOL
VAR_INPUT
	ITFALARM : IAlarm3;
END_VAR
END_METHOD

METHOD MATCHESFILTERCRITERIA2 : BOOL
VAR_INPUT
	ITFALARMMETAOBJECTSTUB5 : IAlarmMetaObjectStub5;
	XCHKPRI : BOOL;
	XCHKGRP : BOOL;
	XCHKCLA : BOOL;
	XCHKLATCH : BOOL;
	XCHKTIMERANGE : BOOL;
END_VAR
END_METHOD

METHOD ELABTIMERANGEFILTERCRITERIA
END_METHOD

METHOD DISPLAYREASONNOTINDEX
END_METHOD

METHOD ELABLATCHFILTERCRITERIA
END_METHOD

METHOD ISLATCHFILTERINDEXABLE : BOOL
VAR_INPUT
	IVERSION : INT;
	EBYTEORDER : EAlarmByteOrder;
	EDBUSED : EDBType;
END_VAR
END_METHOD

METHOD AREALLALARMCLASSESSELECTED : BOOL
END_METHOD

METHOD AREALLALARMGROUPSSELECTED : BOOL
END_METHOD

METHOD GETALARMCLASSES : POINTER TO ARRAY [0..0] OF UDINT
END_METHOD

METHOD GETALARMGROUPS : POINTER TO ARRAY [0..0] OF UDINT
END_METHOD

METHOD GETCOUNTALARMCLASSES : INT
END_METHOD

METHOD GETCOUNTALARMGROUPS : INT
END_METHOD

METHOD GETPRIORITYFROM : USINT
END_METHOD

METHOD GETPRIORITYTO : USINT
END_METHOD

METHOD GETFILTERLATCHCONTENT : INT
END_METHOD

METHOD GETFILTERLATCHTYPEDLITERALTYPE : INT
END_METHOD

METHOD GETFILTERLATCHVALUELI : LINT
END_METHOD

METHOD GETFILTERLATCHVALUELREAL : LREAL
END_METHOD

METHOD GETFILTERLATCHVALUEREAL : REAL
END_METHOD

METHOD GETFILTERLATCHVALUEWSTRING : WSTRING
END_METHOD

METHOD ISFILTERLATCHAVAILABLE : BOOL
END_METHOD

METHOD GETALARMCLASSES3
VAR_OUTPUT
	PASTRUCTFILTERING : POINTER TO ARRAY [0..0] OF StructFilteringName;
	ICOUNT : INT;
END_VAR
END_METHOD

METHOD GETALARMGROUPS3
VAR_OUTPUT
	PASTRUCTFILTERING : POINTER TO ARRAY [0..0] OF StructFilteringName;
	ICOUNT : INT;
END_VAR
END_METHOD

METHOD GETFILTERTIMERANGEFROMVALUELI : LINT
END_METHOD

METHOD GETFILTERTIMERANGETOVALUELI : LINT
END_METHOD

METHOD GETFILTERTIMERANGETYPE : INT
END_METHOD

METHOD ISFILTERTIMERANGEAVAILABLE : BOOL
END_METHOD

METHOD PRVCALCCHECKSUM : WORD
VAR_INPUT
	PDATA : POINTER TO ARRAY [0..0] OF BYTE;
	ISIZE : INT;
END_VAR
END_METHOD

METHOD PRVCHECKSUMFORVARIATION : WORD
END_METHOD

METHOD PRVGETLIVALUE : BOOL
VAR_INPUT
	PVALUE : POINTER TO BYTE;
	EVARIABLETYPE : Visu_Types;
END_VAR
VAR_OUTPUT
	LIVALUE : LINT;
	PDEBUG : POINTER TO ARRAY [0..7] OF BYTE;
END_VAR
END_METHOD

METHOD PRVISCONSIDEREDASNUMERICTYPE : BOOL
VAR_INPUT
	EVARIABLETYPE : Visu_Types;
END_VAR
END_METHOD

METHOD PRVREADLATCHVARVALUE : STO.ERROR
VAR_INPUT
	ITFDATABASEACCESS : IDatabaseAccess;
	USIWHICHLATCHVAR : USINT;
	SVARVALUE : REFERENCE TO STRING;
	SZSVARVALUE : CAA.SIZE;
	WSVARVALUE : REFERENCE TO WSTRING;
	SZWSVARVALUE : CAA.SIZE;
END_VAR
VAR_OUTPUT
	XNULL : BOOL;
	BYTYPE : BYTE;
	LIVALUE : LINT;
END_VAR
END_METHOD

METHOD PRVSWAPBYTES
VAR_INPUT
	PBAVALUE : POINTER TO ARRAY [0..7] OF BYTE;
	IINDEX1 : INT;
	IINDEX2 : INT;
END_VAR
END_METHOD

METHOD PRVSWAPLIVALUE : BOOL
VAR_INPUT
	LIVALUEINP : LINT;
	THETYPE : __SYSTEM.TYPE_CLASS;
END_VAR
VAR_OUTPUT
	LIVALUEOUT : LINT;
END_VAR
END_METHOD

METHOD PRVMATCHESFILTERCRITERIACLASS : BOOL
VAR_INPUT
	UDIALARMCLASSID : UDINT;
	XREMOTEALM : BOOL;
	SPROXYNAME : STRING;
END_VAR
END_METHOD

METHOD PRVMATCHESFILTERCRITERIAGROUPS : BOOL
VAR_INPUT
	UDIALARMGROUPID : UDINT;
	XREMOTEALM : BOOL;
	SPROXYNAME : STRING;
END_VAR
END_METHOD

METHOD PRVMATCHESFILTERCRITERIALATCHVAR : BOOL
VAR_INPUT
	LATCHTYPEDVALUE : ITypedValue;
END_VAR
END_METHOD

METHOD PRVMATCHESFILTERCRITERIAPRIORITY : BOOL
VAR_INPUT
	USIPRIORITY : USINT;
END_VAR
END_METHOD

METHOD PRVMATCHESFILTERCRITERIATIMERANGE : BOOL
VAR_INPUT
	TSTAMPLAST : Timestamp;
	TSTAMPACTIVE : Timestamp;
END_VAR
END_METHOD

(* ---- VISUFBALARMFILTERCRITERIASERVICE.pou ---- *)
FUNCTION_BLOCK VISUFBALARMFILTERCRITERIASERVICE EXTENDS VisuFbAlarmFilterCriteria
END_FUNCTION_BLOCK

METHOD ELABLATCHFILTERCRITERIA
END_METHOD

METHOD ELABTIMERANGEFILTERCRITERIA
END_METHOD

METHOD ISFILTERLATCHAVAILABLE : BOOL
END_METHOD

METHOD ISFILTERTIMERANGEAVAILABLE : BOOL
END_METHOD

(* ---- VISUFBALARMFILTERCRITERIAUSERCLIENT.pou ---- *)
FUNCTION_BLOCK VISUFBALARMFILTERCRITERIAUSERCLIENT EXTENDS VisuFbAlarmFilterCriteria
VAR
	M_AGROUPIDS : ARRAY [0..MAX_ID] OF UDINT;
	M_ACLASSIDS : ARRAY [0..MAX_ID] OF UDINT;
	M_PACLASSIDS : POINTER TO ARRAY [0..0] OF UDINT;
	M_PAGROUPIDS : POINTER TO ARRAY [0..0] OF UDINT;
	M_AGROUPIDSREM : ARRAY [0..MAX_ID] OF StruFilterRemoteAlm;
	M_ACLASSIDSREM : ARRAY [0..MAX_ID] OF StruFilterRemoteAlm;
	M_PACLASSIDSREM : POINTER TO ARRAY [0..0] OF StruFilterRemoteAlm;
	M_PAGROUPIDSREM : POINTER TO ARRAY [0..0] OF StruFilterRemoteAlm;
	MAX_ID : INT := 20;
END_VAR
END_FUNCTION_BLOCK

METHOD ELABLATCHFILTERCRITERIA
END_METHOD

METHOD ELABTIMERANGEFILTERCRITERIA
END_METHOD

METHOD FB_EXIT : BOOL
VAR_INPUT
	BINCOPYCODE : BOOL;
END_VAR
END_METHOD

METHOD INITIALIZE
VAR_INPUT
	ITFALARMFILTERCRITERIA : IAlarmFilterCriteria;
END_VAR
END_METHOD

METHOD ISFILTERLATCHAVAILABLE : BOOL
END_METHOD

METHOD GETALARMCLASSES3
VAR_OUTPUT
	PASTRUCTFILTERING : POINTER TO ARRAY [0..0] OF StructFilteringName;
	ICOUNT : INT;
END_VAR
END_METHOD

METHOD GETALARMGROUPS3
VAR_OUTPUT
	PASTRUCTFILTERING : POINTER TO ARRAY [0..0] OF StructFilteringName;
	ICOUNT : INT;
END_VAR
END_METHOD

METHOD ISFILTERTIMERANGEAVAILABLE : BOOL
END_METHOD
